Fanuc KAREL source: kc00033.KL

-- PROVISIONAL review KL for V1013-1; original PC SHA256 9e4ed1c71de85553b20a89be951cd6529a8f0dabc5021b035f0b5729e391d0ed
-- Incomplete behavior may be omitted. Consult companion uncertainty JSON. Do not deploy.
PROGRAM KC00033
%NOLOCKGROUP
BEGIN
  -- UNRESOLVED_PC offsets 5-32; opcodes 27,22,1C,22,22,76
  -- UNRESOLVED_PC offsets 37-41; opcodes 7F
END KC00033
